TYPE E_BuzzerMode :
(
	eBuzzerOff := 0,
	eBuzzerError,		//Short Delay Off
	eBuzzerWarning		//Long Delay Off
);
END_TYPE

(* stored: Version 1.1.0.1, ProductVersion 3.1.4024.13
   DUT E_BuzzerMode: Id {de52cb38-8c30-4811-9aac-efd92215c3d4} *)
